# EPICS substitutions: db/Beckhoff_7XXX/ecmcEX72XX_OPT_followingError.substitutions
file "ecmc_analogInput-chX.template"
{
  pattern {CH_ID, sourceName, KEY, suffix, DESC, EGU, ESLO, PREC, LOPR, HOPR, LOLO, LOW, HIGH, HIHI, HYST, LLSV, LSV, HSV, HHSV}
          {"$(OPT_CH_ID=01)", "followingError", "Drv", "-PosDiff", "Following Error", "Cnts", 1, 0, 0, 0, 0, 0, 0, 0, 0, "NO_ALARM", "NO_ALARM", "NO_ALARM", "NO_ALARM"}
}
